(* IEC 61131-3 sources: plc-st-coding-agent/progress/evidence/f14_v10_full_20261113/jobs/custom_deepseek-v4pro (part 5) *)

(* ---- self-hard-02.candidate_02.st ---- *)
(* ENGINEERING_CONTRACT
   - Outputs: phase, elapsed, timeout; initial (0,0,FALSE).
   - Priority: abort > new start edge > run counting (PUB002-006).
   - abortBtn TRUE: phase=9, elapsed/timeout hold previous values. Start edge consumed (PUB003, PUB005-006).
   - New start edge without abort: phase=1, elapsed=0, timeout=FALSE; start scan not counted (PUB004, PUB006).
   - Previous scan running (1 or 2), no abort, no start edge: increment elapsed by 1.
     If elapsed >= maxDuration: timeout=TRUE, phase=3 (timeout priority). Else phase=2 if pv>=setpoint or prevPhase=2, otherwise phase=1 (PUB005-006).
   - Phase 3 complete, phase 9 aborted: freeze elapsed, timeout, phase until new valid start or abort.
   - Unit: elapsed counts scans; maxDuration positive integer scan threshold; comparison >=.
*)
FUNCTION_BLOCK FB
VAR_INPUT
    startBtn : BOOL;
    abortBtn : BOOL;
    setpoint : REAL;
    pv : REAL;
    maxDuration : INT;
END_VAR
VAR_OUTPUT
    elapsed : INT;
    phase : INT;
    timeout : BOOL;
END_VAR
VAR
    prevStartBtn : BOOL := FALSE;
    prevPhase : INT := 0;
    prevElapsed : INT := 0;
    prevTimeout : BOOL := FALSE;
    startEdge : BOOL;
END_VAR

(* Record startBtn rising edge before priority processing; consumed even if abort *)
startEdge := startBtn AND NOT prevStartBtn;

IF abortBtn THEN
    (* Abort highest priority: enter phase 9 and freeze elapsed/timeout *)
    phase := 9;
    elapsed := prevElapsed;
    timeout := prevTimeout;
ELSIF startEdge THEN
    (* New valid start with no abort: reset batch and do not count this scan *)
    phase := 1;
    elapsed := 0;
    timeout := FALSE;
ELSE
    (* No abort and no new start edge *)
    IF (prevPhase = 1) OR (prevPhase = 2) THEN
        (* Running state: count exactly one scan *)
        elapsed := prevElapsed + 1;

        IF elapsed >= maxDuration THEN
            (* Timeout has priority over temperature threshold *)
            timeout := TRUE;
            phase := 3;
        ELSE
            timeout := FALSE;
            IF (prevPhase = 2) OR (pv >= setpoint) THEN
                phase := 2;
            ELSE
                phase := 1;
            END_IF;
        END_IF;
    ELSE
        (* Idle, complete, or aborted: hold state *)
        phase := prevPhase;
        elapsed := prevElapsed;
        timeout := prevTimeout;
    END_IF;
END_IF;

(* Update previous-cycle memory *)
prevStartBtn := startBtn;
prevPhase := phase;
prevElapsed := elapsed;
prevTimeout := timeout;

(* CONTRACT_RULES [] *)
END_FUNCTION_BLOCK

(* ---- self-hard-02.raw_candidate_01.st ---- *)
(* ENGINEERING_CONTRACT
   - phase: 0 idle initial; new start & !abort -> 1; in running, elapsed<maxDuration and (prevPhase=2 or pv>=setpoint) -> 2, else 1; elapsed>=maxDuration -> 3; abort -> 9. Priority abort > start edge > run count (PUB002-006).
   - elapsed: increment exactly once per scan when !abort, !startEdge, prevPhase=1/2; reset 0 on new start; freeze otherwise.
   - timeout: set TRUE exactly when running scan counted reaches maxDuration; reset FALSE on new start; freeze on abort/completion/idle.
   - start rising edge recorded first and consumed even if abort same scan; restart requires release/press.
   - maxDuration positive scan count; comparison >=. Boundaries: counts scan after start not counted.
*)
FUNCTION_BLOCK FB
VAR
    prevStartBtn : BOOL := FALSE;
    prevPhase : INT := 0;
    prevElapsed : INT := 0;
    prevTimeout : BOOL := FALSE;
    startEdge : BOOL;
END_VAR

(* Record startBtn rising edge before priority processing; consumed even if abort *)
startEdge := startBtn AND NOT prevStartBtn;

IF abortBtn THEN
    (* Abort has highest priority: enter phase 9 and freeze elapsed/timeout *)
    phase := 9;
    elapsed := prevElapsed;
    timeout := prevTimeout;
ELSIF startEdge THEN
    (* New valid start with no abort: reset batch and do not count this scan *)
    phase := 1;
    elapsed := 0;
    timeout := FALSE;
ELSE
    (* No abort and no new start edge *)
    IF (prevPhase = 1) OR (prevPhase = 2) THEN
        (* Running state: count exactly one scan *)
        elapsed := prevElapsed + 1;

        IF elapsed >= maxDuration THEN
            (* Timeout has priority over temperature threshold *)
            timeout := TRUE;
            phase := 3;
        ELSE
            timeout := FALSE;
            IF (prevPhase = 2) OR (pv >= setpoint) THEN
                phase := 2;
            ELSE
                phase := 1;
            END_IF;
        END_IF;
    ELSE
        (* Idle, complete, or aborted: hold state *)
        phase := prevPhase;
        elapsed := prevElapsed;
        timeout := prevTimeout;
    END_IF;
END_IF;

(* Update previous-cycle memory *)
prevStartBtn := startBtn;
prevPhase := phase;
prevElapsed := elapsed;
prevTimeout := timeout;

(* CONTRACT_RULES [] *)
END_FUNCTION_BLOCK

(* ---- self-hard-02.raw_candidate_02.st ---- *)
(* ENGINEERING_CONTRACT
   - Outputs: phase, elapsed, timeout; initial (0,0,FALSE).
   - Priority: abort > new start edge > run counting (PUB002-006).
   - abortBtn TRUE: phase=9, elapsed/timeout hold previous values. Start edge consumed (PUB003, PUB005-006).
   - New start edge without abort: phase=1, elapsed=0, timeout=FALSE; start scan not counted (PUB004, PUB006).
   - Previous scan running (1 or 2), no abort, no start edge: increment elapsed by 1.
     If elapsed >= maxDuration: timeout=TRUE, phase=3 (timeout priority). Else phase=2 if pv>=setpoint or prevPhase=2, otherwise phase=1 (PUB005-006).
   - Phase 3 complete, phase 9 aborted: freeze elapsed, timeout, phase until new valid start or abort.
   - Unit: elapsed counts scans; maxDuration positive integer scan threshold; comparison >=.
*)
FUNCTION_BLOCK FB
VAR_INPUT
    startBtn : BOOL;
    abortBtn : BOOL;
    setpoint : REAL;
    pv : REAL;
    maxDuration : INT;
END_VAR
VAR_OUTPUT
    elapsed : INT;
    phase : INT;
    timeout : BOOL;
END_VAR
VAR
    prevStartBtn : BOOL := FALSE;
    prevPhase : INT := 0;
    prevElapsed : INT := 0;
    prevTimeout : BOOL := FALSE;
    startEdge : BOOL;
END_VAR

(* Record startBtn rising edge before priority processing; consumed even if abort *)
startEdge := startBtn AND NOT prevStartBtn;

IF abortBtn THEN
    (* Abort highest priority: enter phase 9 and freeze elapsed/timeout *)
    phase := 9;
    elapsed := prevElapsed;
    timeout := prevTimeout;
ELSIF startEdge THEN
    (* New valid start with no abort: reset batch and do not count this scan *)
    phase := 1;
    elapsed := 0;
    timeout := FALSE;
ELSE
    (* No abort and no new start edge *)
    IF (prevPhase = 1) OR (prevPhase = 2) THEN
        (* Running state: count exactly one scan *)
        elapsed := prevElapsed + 1;

        IF elapsed >= maxDuration THEN
            (* Timeout has priority over temperature threshold *)
            timeout := TRUE;
            phase := 3;
        ELSE
            timeout := FALSE;
            IF (prevPhase = 2) OR (pv >= setpoint) THEN
                phase := 2;
            ELSE
                phase := 1;
            END_IF;
        END_IF;
    ELSE
        (* Idle, complete, or aborted: hold state *)
        phase := prevPhase;
        elapsed := prevElapsed;
        timeout := prevTimeout;
    END_IF;
END_IF;

(* Update previous-cycle memory *)
prevStartBtn := startBtn;
prevPhase := phase;
prevElapsed := elapsed;
prevTimeout := timeout;

(* CONTRACT_RULES [] *)
END_FUNCTION_BLOCK

(* ---- self-hard-03.candidate_01.st ---- *)
(* ENGINEERING_CONTRACT
   Activation: pushEn/popEn rising edges vs stored previous inputs; no repeat while held (PUB001-PUB039).
   Same-scan priority: pop edge is processed first, then push edge; simultaneous full pair frees a slot then appends; simultaneous empty pair adds only new item (PUB001-PUB039).
   Retention: tmp_count is static queue length; fifo[1..tmp_count] stays compact on each scan. No explicit reset; only successful edge actions alter valid queue state (PUB001-PUB039).
   Outputs: count := tmp_count; full := tmp_count = 8; empty := tmp_count = 0; head := fifo[1] when nonempty, else 0 (PUB001-PUB039).
   Bounds: count/INT 0..8; fifo indices 1..8. Invalid tail fifo[tmp_count+1..8] is unspecified and not cleared (PUB001-PUB039).
*)
(* CONTRACT_RULES [] *)
FUNCTION_BLOCK FB
VAR_INPUT
    pushEn : BOOL;
    pushItem : INT;
    popEn : BOOL;
END_VAR
VAR_IN_OUT
    fifo : ARRAY[1..8] OF INT;
END_VAR
VAR_OUTPUT
    count : INT;
    full : BOOL;
    empty : BOOL;
    head : INT;
END_VAR
VAR
    prevPushEn : BOOL := FALSE;
    prevPopEn : BOOL := FALSE;
    tmp_count : INT := 0;
    tmp_pushRise : BOOL;
    tmp_popRise : BOOL;
    tmp_i : INT;
END_VAR

tmp_pushRise := pushEn AND NOT prevPushEn;
tmp_popRise := popEn AND NOT prevPopEn;

IF tmp_popRise THEN
    IF tmp_count > 0 THEN
        IF tmp_count > 1 THEN
            FOR tmp_i := 1 TO tmp_count - 1 DO
                fifo[tmp_i] := fifo[tmp_i + 1];
            END_FOR;
        END_IF;
        tmp_count := tmp_count - 1;
    END_IF;
END_IF;

IF tmp_pushRise THEN
    IF tmp_count < 8 THEN
        tmp_count := tmp_count + 1;
        fifo[tmp_count] := pushItem;
    END_IF;
END_IF;

count := tmp_count;
full := (tmp_count = 8);
empty := (tmp_count = 0);

IF tmp_count > 0 THEN
    head := fifo[1];
ELSE
    head := 0;
END_IF;

prevPushEn := pushEn;
prevPopEn := popEn;

END_FUNCTION_BLOCK

(* ---- self-hard-03.raw_candidate_01.st ---- *)
(* ENGINEERING_CONTRACT
   Activation: pushEn/popEn rising edges vs stored previous inputs; no repeat while held (PUB001-PUB039).
   Same-scan priority: pop edge is processed first, then push edge; simultaneous full pair frees a slot then appends; simultaneous empty pair adds only new item (PUB001-PUB039).
   Retention: tmp_count is static queue length; fifo[1..tmp_count] stays compact on each scan. No explicit reset; only successful edge actions alter valid queue state (PUB001-PUB039).
   Outputs: count := tmp_count; full := tmp_count = 8; empty := tmp_count = 0; head := fifo[1] when nonempty, else 0 (PUB001-PUB039).
   Bounds: count/INT 0..8; fifo indices 1..8. Invalid tail fifo[tmp_count+1..8] is unspecified and not cleared (PUB001-PUB039).
*)
(* CONTRACT_RULES [] *)
FUNCTION_BLOCK FB
VAR_INPUT
    pushEn : BOOL;
    pushItem : INT;
    popEn : BOOL;
END_VAR
VAR_IN_OUT
    fifo : ARRAY[1..8] OF INT;
END_VAR
VAR_OUTPUT
    count : INT;
    full : BOOL;
    empty : BOOL;
    head : INT;
END_VAR
VAR
    prevPushEn : BOOL := FALSE;
    prevPopEn : BOOL := FALSE;
    tmp_count : INT := 0;
    tmp_pushRise : BOOL;
    tmp_popRise : BOOL;
    tmp_i : INT;
END_VAR

tmp_pushRise := pushEn AND NOT prevPushEn;
tmp_popRise := popEn AND NOT prevPopEn;

IF tmp_popRise THEN
    IF tmp_count > 0 THEN
        IF tmp_count > 1 THEN
            FOR tmp_i := 1 TO tmp_count - 1 DO
                fifo[tmp_i] := fifo[tmp_i + 1];
            END_FOR;
        END_IF;
        tmp_count := tmp_count - 1;
    END_IF;
END_IF;

IF tmp_pushRise THEN
    IF tmp_count < 8 THEN
        tmp_count := tmp_count + 1;
        fifo[tmp_count] := pushItem;
    END_IF;
END_IF;

count := tmp_count;
full := (tmp_count = 8);
empty := (tmp_count = 0);

IF tmp_count > 0 THEN
    head := fifo[1];
ELSE
    head := 0;
END_IF;

prevPushEn := pushEn;
prevPopEn := popEn;

END_FUNCTION_BLOCK

(* ---- self-hard-05.candidate_01.st ---- *)
(* ENGINEERING_CONTRACT
   tripLatched: set same-scan on runRequest AND NOT flameOK; held until reset rising edge
                with runRequest=FALSE AND flameOK=FALSE only. Same-scan set/reset mutually exclusive.
   fuelPermit : runRequest AND flameOK AND NOT tripLatched; computed after trip update.
   trimEnable : fuelPermit AND NOT o2Fault.
   airTrim    : trimEnable ? clamp(2.0*(2.0-o2PV), -10.0, 10.0) : 0.0; REAL percent.
   airCommand : fuelPermit ? clamp(baseAir+airTrim, 0.0, 100.0) : 0.0; REAL percent.
   o2Fault    : NOT o2Valid OR o2PV<0.0 OR o2PV>21.0; combinational.
*)
(* CONTRACT_RULES [] *)
FUNCTION_BLOCK FB
VAR_INPUT
    runRequest : BOOL;
    flameOK    : BOOL;
    o2Valid    : BOOL;
    o2PV       : REAL;
    baseAir    : REAL;
    resetBtn   : BOOL;
END_VAR
VAR_OUTPUT
    fuelPermit  : BOOL;
    trimEnable  : BOOL;
    airTrim     : REAL;
    airCommand  : REAL;
    tripLatched : BOOL;
    o2Fault     : BOOL;
END_VAR
VAR
    fbResetEdge     : R_TRIG;
    tmp_resetRising : BOOL;
    tmp_trim        : REAL;
    tmp_cmd         : REAL;
END_VAR

fbResetEdge(CLK := resetBtn);
tmp_resetRising := fbResetEdge.Q;

(* Trip latch: same-scan loss-of-flame set; only valid safe-state reset edge clears. *)
tripLatched := (runRequest AND NOT flameOK)
               OR (tripLatched AND NOT (tmp_resetRising AND NOT runRequest AND NOT flameOK));

(* Oxygen analyzer fault and permits. *)
o2Fault := (NOT o2Valid) OR (o2PV < 0.0) OR (o2PV > 21.0);
fuelPermit := runRequest AND flameOK AND NOT tripLatched;
trimEnable := fuelPermit AND NOT o2Fault;

(* Oxygen trim with +/-10 percent output clamp. *)
IF trimEnable THEN
    tmp_trim := 2.0 * (2.0 - o2PV);
    IF tmp_trim < -10.0 THEN
        tmp_trim := -10.0;
    ELSIF tmp_trim > 10.0 THEN
        tmp_trim := 10.0;
    END_IF;
    airTrim := tmp_trim;
ELSE
    airTrim := 0.0;
END_IF;

(* Final air command with 0..100 percent output clamp. *)
IF fuelPermit THEN
    tmp_cmd := baseAir + airTrim;
    IF tmp_cmd < 0.0 THEN
        tmp_cmd := 0.0;
    ELSIF tmp_cmd > 100.0 THEN
        tmp_cmd := 100.0;
    END_IF;
    airCommand := tmp_cmd;
ELSE
    airCommand := 0.0;
END_IF;

END_FUNCTION_BLOCK

(* ---- self-hard-05.raw_candidate_01.st ---- *)
(* ENGINEERING_CONTRACT
   tripLatched: set same-scan on runRequest AND NOT flameOK; held until reset rising edge
                with runRequest=FALSE AND flameOK=FALSE only. Same-scan set/reset mutually exclusive.
   fuelPermit : runRequest AND flameOK AND NOT tripLatched; computed after trip update.
   trimEnable : fuelPermit AND NOT o2Fault.
   airTrim    : trimEnable ? clamp(2.0*(2.0-o2PV), -10.0, 10.0) : 0.0; REAL percent.
   airCommand : fuelPermit ? clamp(baseAir+airTrim, 0.0, 100.0) : 0.0; REAL percent.
   o2Fault    : NOT o2Valid OR o2PV<0.0 OR o2PV>21.0; combinational.
*)
(* CONTRACT_RULES [] *)
FUNCTION_BLOCK FB
VAR_INPUT
    runRequest : BOOL;
    flameOK    : BOOL;
    o2Valid    : BOOL;
    o2PV       : REAL;
    baseAir    : REAL;
    resetBtn   : BOOL;
END_VAR
VAR_OUTPUT
    fuelPermit  : BOOL;
    trimEnable  : BOOL;
    airTrim     : REAL;
    airCommand  : REAL;
    tripLatched : BOOL;
    o2Fault     : BOOL;
END_VAR
VAR
    fbResetEdge     : R_TRIG;
    tmp_resetRising : BOOL;
    tmp_trim        : REAL;
    tmp_cmd         : REAL;
END_VAR

fbResetEdge(CLK := resetBtn);
tmp_resetRising := fbResetEdge.Q;

(* Trip latch: same-scan loss-of-flame set; only valid safe-state reset edge clears. *)
tripLatched := (runRequest AND NOT flameOK)
               OR (tripLatched AND NOT (tmp_resetRising AND NOT runRequest AND NOT flameOK));

(* Oxygen analyzer fault and permits. *)
o2Fault := (NOT o2Valid) OR (o2PV < 0.0) OR (o2PV > 21.0);
fuelPermit := runRequest AND flameOK AND NOT tripLatched;
trimEnable := fuelPermit AND NOT o2Fault;

(* Oxygen trim with +/-10 percent output clamp. *)
IF trimEnable THEN
    tmp_trim := 2.0 * (2.0 - o2PV);
    IF tmp_trim < -10.0 THEN
        tmp_trim := -10.0;
    ELSIF tmp_trim > 10.0 THEN
        tmp_trim := 10.0;
    END_IF;
    airTrim := tmp_trim;
ELSE
    airTrim := 0.0;
END_IF;

(* Final air command with 0..100 percent output clamp. *)
IF fuelPermit THEN
    tmp_cmd := baseAir + airTrim;
    IF tmp_cmd < 0.0 THEN
        tmp_cmd := 0.0;
    ELSIF tmp_cmd > 100.0 THEN
        tmp_cmd := 100.0;
    END_IF;
    airCommand := tmp_cmd;
ELSE
    airCommand := 0.0;
END_IF;

END_FUNCTION_BLOCK

(* ---- self-hard-06.candidate_01.st ---- *)
(* ENGINEERING_CONTRACT
   - tripLatched: set same scan by run & (!valid | P>=4500) PUB002/PUB006; holds until legal reset edge.
     Legal reset: rising reset & !run & valid & P<=4200 PUB003. Illegal reset does not clear PUB012/PUB013.
   - currentCauseMask: recomputed each scan; allowed 0/1/2/4/6/8 PUB008,N10-S15.
     bit0=invalid; bit1 requires 3 consecutive full stuck scans PUB010,N10-S11; bit2 inclusive flow; bit3=8 when no located bit under overpressure.
   - latchedCauseMask: OR-accumulates currentCauseMask while tripLatched true; cleared when not tripped or legal reset PUB011,N10-S18.
   - fuelPermit = run & !trip; diagnosticActive = current<>0 PUB007.
   - stuck counter zeroes on any non-full scan: !run, !valid, P<4500, or valve condition false PUB010.
   - units: kPa, t/h, %; boundaries inclusive. Same-scan trip and cause are emitted together.
*)
(* CONTRACT_RULES [] *)
FUNCTION_BLOCK FB
VAR_INPUT
    runRequest: BOOL;
    pressure: REAL;
    pressureValid: BOOL;
    fuelFlow: REAL;
    steamFlow: REAL;
    outletCmd: INT;
    outletFeedback: INT;
    resetBtn: BOOL;
END_VAR
VAR_OUTPUT
    tripLatched: BOOL;
    fuelPermit: BOOL;
    currentCauseMask: WORD;
    latchedCauseMask: WORD;
    diagnosticActive: BOOL;
END_VAR
VAR
    prev_reset_btn: BOOL := FALSE;
    prev_trip_state: BOOL := FALSE;
    stuck_count: INT := 0;
    latched_state: WORD := WORD#16#0000;
    tmp_rising_reset: BOOL;
    tmp_legal_reset: BOOL;
    tmp_stuck_condition: BOOL;
    tmp_bit1: BOOL;
    tmp_bit2: BOOL;
    tmp_trip_condition: BOOL;
    tmp_trip_state: BOOL;
END_VAR

(* Update stuck-valve consecutive-scan counter *)
tmp_stuck_condition := runRequest AND pressureValid AND (pressure >= 4500.0)
                       AND (outletCmd >= 50) AND (outletFeedback <= 10);

IF tmp_stuck_condition THEN
    IF stuck_count < 3 THEN
        stuck_count := stuck_count + 1;
    END_IF;
ELSE
    stuck_count := 0;
END_IF;

(* Compute current cause mask *)
currentCauseMask := WORD#16#0000;

IF NOT runRequest THEN
    currentCauseMask := WORD#16#0000;
ELSIF NOT pressureValid THEN
    currentCauseMask := WORD#16#0001; (* bit0: transmitter invalid *)
ELSE
    IF pressure >= 4500.0 THEN
        tmp_bit1 := stuck_count >= 3;
        tmp_bit2 := (fuelFlow >= 4.0) AND (steamFlow <= 10.0);

        IF tmp_bit1 THEN
            currentCauseMask := currentCauseMask OR WORD#16#0002; (* bit1: valve stuck *)
        END_IF;
        IF tmp_bit2 THEN
            currentCauseMask := currentCauseMask OR WORD#16#0004; (* bit2: combustion excess *)
        END_IF;
        IF currentCauseMask = WORD#16#0000 THEN
            currentCauseMask := WORD#16#0008; (* bit3: not located *)
        END_IF;
    ELSE
        currentCauseMask := WORD#16#0000;
    END_IF;
END_IF;

(* Trip latch state *)
tmp_rising_reset := resetBtn AND NOT prev_reset_btn;
tmp_legal_reset := tmp_rising_reset AND (NOT runRequest) AND pressureValid AND (pressure <= 4200.0);

tmp_trip_condition := runRequest AND ((NOT pressureValid) OR (pressureValid AND (pressure >= 4500.0)));
tmp_trip_state := tmp_trip_condition OR (prev_trip_state AND NOT tmp_legal_reset);
tripLatched := tmp_trip_state;

(* Latched footprint accumulation / clear *)
IF tmp_trip_state THEN
    latched_state := (latched_state OR currentCauseMask) AND WORD#16#000F;
ELSE
    latched_state := WORD#16#0000;
END_IF;
latchedCauseMask := latched_state;

(* Derived outputs *)
fuelPermit := runRequest AND NOT tripLatched;
diagnosticActive := currentCauseMask <> WORD#16#0000;

(* Remember previous-scan values for next call *)
prev_reset_btn := resetBtn;
prev_trip_state := tmp_trip_state;

END_FUNCTION_BLOCK

(* ---- self-hard-06.raw_candidate_01.st ---- *)
(* ENGINEERING_CONTRACT
   - tripLatched: set same scan by run & (!valid | P>=4500) PUB002/PUB006; holds until legal reset edge.
     Legal reset: rising reset & !run & valid & P<=4200 PUB003. Illegal reset does not clear PUB012/PUB013.
   - currentCauseMask: recomputed each scan; allowed 0/1/2/4/6/8 PUB008,N10-S15.
     bit0=invalid; bit1 requires 3 consecutive full stuck scans PUB010,N10-S11; bit2 inclusive flow; bit3=8 when no located bit under overpressure.
   - latchedCauseMask: OR-accumulates currentCauseMask while tripLatched true; cleared when not tripped or legal reset PUB011,N10-S18.
   - fuelPermit = run & !trip; diagnosticActive = current<>0 PUB007.
   - stuck counter zeroes on any non-full scan: !run, !valid, P<4500, or valve condition false PUB010.
   - units: kPa, t/h, %; boundaries inclusive. Same-scan trip and cause are emitted together.
*)
(* CONTRACT_RULES [] *)
FUNCTION_BLOCK FB
VAR_INPUT
    runRequest: BOOL;
    pressure: REAL;
    pressureValid: BOOL;
    fuelFlow: REAL;
    steamFlow: REAL;
    outletCmd: INT;
    outletFeedback: INT;
    resetBtn: BOOL;
END_VAR
VAR_OUTPUT
    tripLatched: BOOL;
    fuelPermit: BOOL;
    currentCauseMask: WORD;
    latchedCauseMask: WORD;
    diagnosticActive: BOOL;
END_VAR
VAR
    prev_reset_btn: BOOL := FALSE;
    prev_trip_state: BOOL := FALSE;
    stuck_count: INT := 0;
    latched_state: WORD := WORD#16#0000;
    tmp_rising_reset: BOOL;
    tmp_legal_reset: BOOL;
    tmp_stuck_condition: BOOL;
    tmp_bit1: BOOL;
    tmp_bit2: BOOL;
    tmp_trip_condition: BOOL;
    tmp_trip_state: BOOL;
END_VAR

(* Update stuck-valve consecutive-scan counter *)
tmp_stuck_condition := runRequest AND pressureValid AND (pressure >= 4500.0)
                       AND (outletCmd >= 50) AND (outletFeedback <= 10);

IF tmp_stuck_condition THEN
    IF stuck_count < 3 THEN
        stuck_count := stuck_count + 1;
    END_IF;
ELSE
    stuck_count := 0;
END_IF;

(* Compute current cause mask *)
currentCauseMask := WORD#16#0000;

IF NOT runRequest THEN
    currentCauseMask := WORD#16#0000;
ELSIF NOT pressureValid THEN
    currentCauseMask := WORD#16#0001; (* bit0: transmitter invalid *)
ELSE
    IF pressure >= 4500.0 THEN
        tmp_bit1 := stuck_count >= 3;
        tmp_bit2 := (fuelFlow >= 4.0) AND (steamFlow <= 10.0);

        IF tmp_bit1 THEN
            currentCauseMask := currentCauseMask OR WORD#16#0002; (* bit1: valve stuck *)
        END_IF;
        IF tmp_bit2 THEN
            currentCauseMask := currentCauseMask OR WORD#16#0004; (* bit2: combustion excess *)
        END_IF;
        IF currentCauseMask = WORD#16#0000 THEN
            currentCauseMask := WORD#16#0008; (* bit3: not located *)
        END_IF;
    ELSE
        currentCauseMask := WORD#16#0000;
    END_IF;
END_IF;

(* Trip latch state *)
tmp_rising_reset := resetBtn AND NOT prev_reset_btn;
tmp_legal_reset := tmp_rising_reset AND (NOT runRequest) AND pressureValid AND (pressure <= 4200.0);

tmp_trip_condition := runRequest AND ((NOT pressureValid) OR (pressureValid AND (pressure >= 4500.0)));
tmp_trip_state := tmp_trip_condition OR (prev_trip_state AND NOT tmp_legal_reset);
tripLatched := tmp_trip_state;

(* Latched footprint accumulation / clear *)
IF tmp_trip_state THEN
    latched_state := (latched_state OR currentCauseMask) AND WORD#16#000F;
ELSE
    latched_state := WORD#16#0000;
END_IF;
latchedCauseMask := latched_state;

(* Derived outputs *)
fuelPermit := runRequest AND NOT tripLatched;
diagnosticActive := currentCauseMask <> WORD#16#0000;

(* Remember previous-scan values for next call *)
prev_reset_btn := resetBtn;
prev_trip_state := tmp_trip_state;

END_FUNCTION_BLOCK

(* ---- self-medium-01.candidate_01.st ---- *)
TYPE ST_Recipe :
STRUCT
    recipeID : INT;
    totalRatio : REAL;
    temperature : REAL;
END_STRUCT
END_TYPE;

(* ENGINEERING_CONTRACT
   valid/loadedID activate only on loadCmd rising edge with running=FALSE (PUB003/PUB007/PUB010).
   Legal slot check 1..8 precedes any array access; out-of-range is not indexed (PUB006/S5).
   Candidate = recipeID<>0 AND totalRatio in [99.0,101.0] AND temperature in [30.0,180.0] (PUB008/N10-S7).
   Accepted invalid edge clears valid=FALSE and loadedID=0; valid edge loads selected recipeID (PUB009/N10-S8/S1).
   running=TRUE overrides any load edge and holds previous valid/loadedID (PUB010/N10-S4/N10-S9).
   No rising edge holds previous outputs (S6/S9).
   Units/bounds: REAL closed intervals; no timing; selSlot dimensionless.
   Conflict note: F13-S1 prose says empty-slot must not change ID, but formal S1/N10-S8/req5 require clear; clear is implemented.
*)

(* CONTRACT_RULES [] *)

FUNCTION_BLOCK FB
VAR_INPUT
    recipe : ARRAY[1..8] OF ST_Recipe;
    selSlot : INT;
    loadCmd : BOOL;
    running : BOOL;
END_VAR
VAR_OUTPUT
    valid : BOOL;
    loadedID : INT;
END_VAR
VAR
    tmp_prevLoadCmd : BOOL := FALSE;
    tmp_validState : BOOL := FALSE;
    tmp_loadedIDState : INT := 0;
    tmp_edge : BOOL;
    tmp_slotLegal : BOOL;
    tmp_candidateValid : BOOL;
    tmp_isNonEmpty : BOOL;
    tmp_ratioOk : BOOL;
    tmp_tempOk : BOOL;
    tmp_recipeId : INT;
    tmp_totalRatio : REAL;
    tmp_temperature : REAL;
END_VAR

tmp_edge := loadCmd AND NOT tmp_prevLoadCmd;

IF (NOT running) AND tmp_edge THEN
    tmp_slotLegal := (selSlot >= 1) AND (selSlot <= 8);
    IF tmp_slotLegal THEN
        tmp_recipeId := recipe[selSlot].recipeID;
        tmp_totalRatio := recipe[selSlot].totalRatio;
        tmp_temperature := recipe[selSlot].temperature;

        tmp_isNonEmpty := (tmp_recipeId <> 0);
        tmp_ratioOk := (tmp_totalRatio >= 99.0) AND (tmp_totalRatio <= 101.0);
        tmp_tempOk := (tmp_temperature >= 30.0) AND (tmp_temperature <= 180.0);
        tmp_candidateValid := tmp_isNonEmpty AND tmp_ratioOk AND tmp_tempOk;

        tmp_validState := tmp_candidateValid;
        IF tmp_candidateValid THEN
            tmp_loadedIDState := tmp_recipeId;
        ELSE
            tmp_loadedIDState := 0;
        END_IF;
    ELSE
        tmp_validState := FALSE;
        tmp_loadedIDState := 0;
    END_IF;
END_IF;

valid := tmp_validState;
loadedID := tmp_loadedIDState;
tmp_prevLoadCmd := loadCmd;

END_FUNCTION_BLOCK

(* ---- self-medium-01.raw_candidate_01.st ---- *)
TYPE ST_Recipe :
STRUCT
    recipeID : INT;
    totalRatio : REAL;
    temperature : REAL;
END_STRUCT
END_TYPE

(* ENGINEERING_CONTRACT
   valid/loadedID activate only on loadCmd rising edge with running=FALSE (PUB003/PUB007/PUB010).
   Legal slot check 1..8 precedes any array access; out-of-range is not indexed (PUB006/S5).
   Candidate = recipeID<>0 AND totalRatio in [99.0,101.0] AND temperature in [30.0,180.0] (PUB008/N10-S7).
   Accepted invalid edge clears valid=FALSE and loadedID=0; valid edge loads selected recipeID (PUB009/N10-S8/S1).
   running=TRUE overrides any load edge and holds previous valid/loadedID (PUB010/N10-S4/N10-S9).
   No rising edge holds previous outputs (S6/S9).
   Units/bounds: REAL closed intervals; no timing; selSlot dimensionless.
   Conflict note: F13-S1 prose says empty-slot must not change ID, but formal S1/N10-S8/req5 require clear; clear is implemented.
*)

(* CONTRACT_RULES [] *)

FUNCTION_BLOCK FB
VAR_INPUT
    recipe : ARRAY[1..8] OF ST_Recipe;
    selSlot : INT;
    loadCmd : BOOL;
    running : BOOL;
END_VAR
VAR_OUTPUT
    valid : BOOL;
    loadedID : INT;
END_VAR
VAR
    tmp_prevLoadCmd : BOOL := FALSE;
    tmp_validState : BOOL := FALSE;
    tmp_loadedIDState : INT := 0;
    tmp_edge : BOOL;
    tmp_slotLegal : BOOL;
    tmp_candidateValid : BOOL;
    tmp_isNonEmpty : BOOL;
    tmp_ratioOk : BOOL;
    tmp_tempOk : BOOL;
    tmp_recipeId : INT;
    tmp_totalRatio : REAL;
    tmp_temperature : REAL;
END_VAR

tmp_edge := loadCmd AND NOT tmp_prevLoadCmd;

IF (NOT running) AND tmp_edge THEN
    tmp_slotLegal := (selSlot >= 1) AND (selSlot <= 8);
    IF tmp_slotLegal THEN
        tmp_recipeId := recipe[selSlot].recipeID;
        tmp_totalRatio := recipe[selSlot].totalRatio;
        tmp_temperature := recipe[selSlot].temperature;

        tmp_isNonEmpty := (tmp_recipeId <> 0);
        tmp_ratioOk := (tmp_totalRatio >= 99.0) AND (tmp_totalRatio <= 101.0);
        tmp_tempOk := (tmp_temperature >= 30.0) AND (tmp_temperature <= 180.0);
        tmp_candidateValid := tmp_isNonEmpty AND tmp_ratioOk AND tmp_tempOk;

        tmp_validState := tmp_candidateValid;
        IF tmp_candidateValid THEN
            tmp_loadedIDState := tmp_recipeId;
        ELSE
            tmp_loadedIDState := 0;
        END_IF;
    ELSE
        tmp_validState := FALSE;
        tmp_loadedIDState := 0;
    END_IF;
END_IF;

valid := tmp_validState;
loadedID := tmp_loadedIDState;
tmp_prevLoadCmd := loadCmd;

END_FUNCTION_BLOCK

(* ---- self-medium-02.candidate_01.st ---- *)
FUNCTION_BLOCK FB
VAR_INPUT
    enable : BOOL;
    rawValue : REAL;
END_VAR
VAR_OUTPUT
    filteredValue : REAL;
    windowFull : BOOL;
    sampleCount : INT;
END_VAR
VAR
    local_data : ARRAY[0..7] OF REAL;
    local_count : INT := 0;
    local_writeIdx : INT := 0;
    local_sum : REAL;
    local_idx : INT;
    local_filtered : REAL := 0.0;
END_VAR

(* ENGINEERING_CONTRACT
  [PUB001-PUB003] enable TRUE: insert rawValue into 8-slot FIFO.
  [PUB004-PUB008] count=min(8,prev+1); unfilled slots ignored.
  [PUB009-PUB012] full: replace oldest slot and rotate write index.
  [PUB013-PUB016] sampleCount=count 0..8; windowFull=(count=8).
  [PUB017-PUB020] enable FALSE: clear history, count=0, full=FALSE,
      filteredValue held from last computation.
  [S1-S7] average over first count slots; boundaries strict; output at end.
*)

(* CONTRACT_RULES [] *)

IF enable THEN
    IF local_count < 8 THEN
        local_data[local_count] := rawValue;
        local_count := local_count + 1;
        local_writeIdx := local_count MOD 8;
    ELSE
        local_data[local_writeIdx] := rawValue;
        local_writeIdx := (local_writeIdx + 1) MOD 8;
    END_IF;

    sampleCount := local_count;
    windowFull := (local_count = 8);

    local_sum := 0.0;
    FOR local_idx := 0 TO local_count - 1 DO
        local_sum := local_sum + local_data[local_idx];
    END_FOR;

    local_filtered := local_sum / INT_TO_REAL(local_count);
    filteredValue := local_filtered;
ELSE
    local_count := 0;
    local_writeIdx := 0;
    sampleCount := 0;
    windowFull := FALSE;

    FOR local_idx := 0 TO 7 DO
        local_data[local_idx] := 0.0;
    END_FOR;

    filteredValue := local_filtered;
END_IF;
END_FUNCTION_BLOCK

(* ---- self-medium-02.raw_candidate_01.st ---- *)
FUNCTION_BLOCK FB
VAR_INPUT
    enable : BOOL;
    rawValue : REAL;
END_VAR
VAR_OUTPUT
    filteredValue : REAL;
    windowFull : BOOL;
    sampleCount : INT;
END_VAR
VAR
    local_data : ARRAY[0..7] OF REAL;
    local_count : INT := 0;
    local_writeIdx : INT := 0;
    local_sum : REAL;
    local_idx : INT;
    local_filtered : REAL := 0.0;
END_VAR

(* ENGINEERING_CONTRACT
  [PUB001-PUB003] enable TRUE: insert rawValue into 8-slot FIFO.
  [PUB004-PUB008] count=min(8,prev+1); unfilled slots ignored.
  [PUB009-PUB012] full: replace oldest slot and rotate write index.
  [PUB013-PUB016] sampleCount=count 0..8; windowFull=(count=8).
  [PUB017-PUB020] enable FALSE: clear history, count=0, full=FALSE,
      filteredValue held from last computation.
  [S1-S7] average over first count slots; boundaries strict; output at end.
*)

(* CONTRACT_RULES [] *)

IF enable THEN
    IF local_count < 8 THEN
        local_data[local_count] := rawValue;
        local_count := local_count + 1;
        local_writeIdx := local_count MOD 8;
    ELSE
        local_data[local_writeIdx] := rawValue;
        local_writeIdx := (local_writeIdx + 1) MOD 8;
    END_IF;

    sampleCount := local_count;
    windowFull := (local_count = 8);

    local_sum := 0.0;
    FOR local_idx := 0 TO local_count - 1 DO
        local_sum := local_sum + local_data[local_idx];
    END_FOR;

    local_filtered := local_sum / INT_TO_REAL(local_count);
    filteredValue := local_filtered;
ELSE
    local_count := 0;
    local_writeIdx := 0;
    sampleCount := 0;
    windowFull := FALSE;

    FOR local_idx := 0 TO 7 DO
        local_data[local_idx] := 0.0;
    END_FOR;

    filteredValue := local_filtered;
END_IF;
END_FUNCTION_BLOCK

(* ---- self-medium-03.candidate_01.st ---- *)
(* ENGINEERING_CONTRACT
   state IDLE/OPENING/CLOSING/FAULT retained in FB; initial IDLE, all previous inputs/outputs FALSE.
   motorUp: activates on IDLE legal open edge, holds while no obstacle and no openLimit; stops at limit/obstacle/fault; mutually exclusive with down.
   motorDown: symmetric close handling, holds while no obstacle and no closeLimit; mutually exclusive with up.
   errorFlag: set by obstacle any scan; latched until bothBTN rising edge and no obstacle; obstacle overrides reset; reset scan motors off, state IDLE.
   prev* memory updated after outputs; BOOL units, initial prev FALSE.
*)
(* CONTRACT_RULES [] *)
FUNCTION_BLOCK FB
VAR
    state : INT := 0; (* 0=IDLE, 1=OPENING, 2=CLOSING, 3=FAULT *)
    prevOpenBtn : BOOL := FALSE;
    prevCloseBtn : BOOL := FALSE;
    prevBothBtn : BOOL := FALSE;
    prevMotorUp : BOOL := FALSE;
    prevMotorDown : BOOL := FALSE;
    prevErrorFlag : BOOL := FALSE;
    prevObstacle : BOOL := FALSE;
    risingOpen : BOOL;
    risingClose : BOOL;
    risingBoth : BOOL;
END_VAR

risingOpen := openBtn AND (NOT prevOpenBtn);
risingClose := closeBtn AND (NOT prevCloseBtn);
risingBoth := (openBtn AND closeBtn) AND (NOT prevBothBtn);

motorUp := (NOT obstacle) AND (NOT openLimit) AND
           (prevMotorUp OR
            ((NOT prevMotorUp) AND (NOT prevMotorDown) AND
             (NOT prevErrorFlag) AND risingOpen AND (NOT closeBtn)));

motorDown := (NOT obstacle) AND (NOT closeLimit) AND
             (prevMotorDown OR
              ((NOT prevMotorUp) AND (NOT prevMotorDown) AND
               (NOT prevErrorFlag) AND risingClose AND (NOT openBtn)));

errorFlag := obstacle OR (prevErrorFlag AND (NOT risingBoth));

IF obstacle THEN
    state := 3;
ELSIF state = 3 THEN
    IF risingBoth THEN
        state := 0;
    ELSE
        state := 3;
    END_IF;
ELSE
    IF motorUp THEN
        state := 1;
    ELSIF motorDown THEN
        state := 2;
    ELSE
        state := 0;
    END_IF;
END_IF;

prevOpenBtn := openBtn;
prevCloseBtn := closeBtn;
prevBothBtn := openBtn AND closeBtn;
prevMotorUp := motorUp;
prevMotorDown := motorDown;
prevErrorFlag := errorFlag;
prevObstacle := obstacle;

END_FUNCTION_BLOCK

(* ---- self-medium-03.candidate_02.st ---- *)
(* ENGINEERING_CONTRACT
   State IDLE/OPENING/CLOSING/FAULT retained in FB; initial IDLE, all previous inputs/outputs FALSE.
   motorUp: activates on IDLE legal open edge, holds while no obstacle and no openLimit; stops at limit/obstacle/fault.
   motorDown: symmetric close handling, holds while no obstacle and no closeLimit.
   errorFlag: set by obstacle any scan; latched until bothBTN rising edge and no obstacle; obstacle overrides reset.
   prev* memory updated after outputs; BOOL units, initial prev FALSE.
*)
(* CONTRACT_RULES [] *)
FUNCTION_BLOCK FB
VAR_INPUT
    openBtn : BOOL;
    closeBtn : BOOL;
    openLimit : BOOL;
    closeLimit : BOOL;
    obstacle : BOOL;
END_VAR
VAR_OUTPUT
    motorUp : BOOL;
    motorDown : BOOL;
    errorFlag : BOOL;
END_VAR
VAR
    state : INT := 0; (* 0=IDLE, 1=OPENING, 2=CLOSING, 3=FAULT *)
    prevOpenBtn : BOOL := FALSE;
    prevCloseBtn : BOOL := FALSE;
    prevBothBtn : BOOL := FALSE;
    prevMotorUp : BOOL := FALSE;
    prevMotorDown : BOOL := FALSE;
    prevErrorFlag : BOOL := FALSE;
    prevObstacle : BOOL := FALSE;
    risingOpen : BOOL;
    risingClose : BOOL;
    risingBoth : BOOL;
END_VAR

risingOpen := openBtn AND (NOT prevOpenBtn);
risingClose := closeBtn AND (NOT prevCloseBtn);
risingBoth := (openBtn AND closeBtn) AND (NOT prevBothBtn);

motorUp := (NOT obstacle) AND (NOT openLimit) AND
           (prevMotorUp OR
            ((NOT prevMotorUp) AND (NOT prevMotorDown) AND
             (NOT prevErrorFlag) AND risingOpen AND (NOT closeBtn)));

motorDown := (NOT obstacle) AND (NOT closeLimit) AND
             (prevMotorDown OR
              ((NOT prevMotorUp) AND (NOT prevMotorDown) AND
               (NOT prevErrorFlag) AND risingClose AND (NOT openBtn)));

errorFlag := obstacle OR (prevErrorFlag AND (NOT risingBoth));

IF obstacle THEN
    state := 3;
ELSIF state = 3 THEN
    IF risingBoth THEN
        state := 0;
    ELSE
        state := 3;
    END_IF;
ELSE
    IF motorUp THEN
        state := 1;
    ELSIF motorDown THEN
        state := 2;
    ELSE
        state := 0;
    END_IF;
END_IF;

prevOpenBtn := openBtn;
prevCloseBtn := closeBtn;
prevBothBtn := openBtn AND closeBtn;
prevMotorUp := motorUp;
prevMotorDown := motorDown;
prevErrorFlag := errorFlag;
prevObstacle := obstacle;

END_FUNCTION_BLOCK

(* ---- self-medium-03.raw_candidate_01.st ---- *)
(* ENGINEERING_CONTRACT
   state IDLE/OPENING/CLOSING/FAULT retained in FB; initial IDLE, all previous inputs/outputs FALSE.
   motorUp: activates on IDLE legal open edge, holds while no obstacle and no openLimit; stops at limit/obstacle/fault; mutually exclusive with down.
   motorDown: symmetric close handling, holds while no obstacle and no closeLimit; mutually exclusive with up.
   errorFlag: set by obstacle any scan; latched until bothBTN rising edge and no obstacle; obstacle overrides reset; reset scan motors off, state IDLE.
   prev* memory updated after outputs; BOOL units, initial prev FALSE.
*)
(* CONTRACT_RULES [] *)
FUNCTION_BLOCK FB
VAR
    state : INT := 0; (* 0=IDLE, 1=OPENING, 2=CLOSING, 3=FAULT *)
    prevOpenBtn : BOOL := FALSE;
    prevCloseBtn : BOOL := FALSE;
    prevBothBtn : BOOL := FALSE;
    prevMotorUp : BOOL := FALSE;
    prevMotorDown : BOOL := FALSE;
    prevErrorFlag : BOOL := FALSE;
    prevObstacle : BOOL := FALSE;
    risingOpen : BOOL;
    risingClose : BOOL;
    risingBoth : BOOL;
END_VAR

risingOpen := openBtn AND (NOT prevOpenBtn);
risingClose := closeBtn AND (NOT prevCloseBtn);
risingBoth := (openBtn AND closeBtn) AND (NOT prevBothBtn);

motorUp := (NOT obstacle) AND (NOT openLimit) AND
           (prevMotorUp OR
            ((NOT prevMotorUp) AND (NOT prevMotorDown) AND
             (NOT prevErrorFlag) AND risingOpen AND (NOT closeBtn)));

motorDown := (NOT obstacle) AND (NOT closeLimit) AND
             (prevMotorDown OR
              ((NOT prevMotorUp) AND (NOT prevMotorDown) AND
               (NOT prevErrorFlag) AND risingClose AND (NOT openBtn)));

errorFlag := obstacle OR (prevErrorFlag AND (NOT risingBoth));

IF obstacle THEN
    state := 3;
ELSIF state = 3 THEN
    IF risingBoth THEN
        state := 0;
    ELSE
        state := 3;
    END_IF;
ELSE
    IF motorUp THEN
        state := 1;
    ELSIF motorDown THEN
        state := 2;
    ELSE
        state := 0;
    END_IF;
END_IF;

prevOpenBtn := openBtn;
prevCloseBtn := closeBtn;
prevBothBtn := openBtn AND closeBtn;
prevMotorUp := motorUp;
prevMotorDown := motorDown;
prevErrorFlag := errorFlag;
prevObstacle := obstacle;

END_FUNCTION_BLOCK

(* ---- self-medium-03.raw_candidate_02.st ---- *)
(* ENGINEERING_CONTRACT
   State IDLE/OPENING/CLOSING/FAULT retained in FB; initial IDLE, all previous inputs/outputs FALSE.
   motorUp: activates on IDLE legal open edge, holds while no obstacle and no openLimit; stops at limit/obstacle/fault.
   motorDown: symmetric close handling, holds while no obstacle and no closeLimit.
   errorFlag: set by obstacle any scan; latched until bothBTN rising edge and no obstacle; obstacle overrides reset.
   prev* memory updated after outputs; BOOL units, initial prev FALSE.
*)
(* CONTRACT_RULES [] *)
FUNCTION_BLOCK FB
VAR_INPUT
    openBtn : BOOL;
    closeBtn : BOOL;
    openLimit : BOOL;
    closeLimit : BOOL;
    obstacle : BOOL;
END_VAR
VAR_OUTPUT
    motorUp : BOOL;
    motorDown : BOOL;
    errorFlag : BOOL;
END_VAR
VAR
    state : INT := 0; (* 0=IDLE, 1=OPENING, 2=CLOSING, 3=FAULT *)
    prevOpenBtn : BOOL := FALSE;
    prevCloseBtn : BOOL := FALSE;
    prevBothBtn : BOOL := FALSE;
    prevMotorUp : BOOL := FALSE;
    prevMotorDown : BOOL := FALSE;
    prevErrorFlag : BOOL := FALSE;
    prevObstacle : BOOL := FALSE;
    risingOpen : BOOL;
    risingClose : BOOL;
    risingBoth : BOOL;
END_VAR

risingOpen := openBtn AND (NOT prevOpenBtn);
risingClose := closeBtn AND (NOT prevCloseBtn);
risingBoth := (openBtn AND closeBtn) AND (NOT prevBothBtn);

motorUp := (NOT obstacle) AND (NOT openLimit) AND
           (prevMotorUp OR
            ((NOT prevMotorUp) AND (NOT prevMotorDown) AND
             (NOT prevErrorFlag) AND risingOpen AND (NOT closeBtn)));

motorDown := (NOT obstacle) AND (NOT closeLimit) AND
             (prevMotorDown OR
              ((NOT prevMotorUp) AND (NOT prevMotorDown) AND
               (NOT prevErrorFlag) AND risingClose AND (NOT openBtn)));

errorFlag := obstacle OR (prevErrorFlag AND (NOT risingBoth));

IF obstacle THEN
    state := 3;
ELSIF state = 3 THEN
    IF risingBoth THEN
        state := 0;
    ELSE
        state := 3;
    END_IF;
ELSE
    IF motorUp THEN
        state := 1;
    ELSIF motorDown THEN
        state := 2;
    ELSE
        state := 0;
    END_IF;
END_IF;

prevOpenBtn := openBtn;
prevCloseBtn := closeBtn;
prevBothBtn := openBtn AND closeBtn;
prevMotorUp := motorUp;
prevMotorDown := motorDown;
prevErrorFlag := errorFlag;
prevObstacle := obstacle;

END_FUNCTION_BLOCK

(* ---- self-medium-04.candidate_01.st ---- *)
FUNCTION_BLOCK FB
VAR_INPUT
    startBtn : BOOL;
    resetBtn : BOOL;
    doneSensor : BOOL;
    targetVol : REAL;
    flowVol : REAL;
END_VAR
VAR_OUTPUT
    valveOpen : BOOL;
    fillsToday : INT;
END_VAR
VAR
    start_prev : BOOL := FALSE;
    reset_prev : BOOL := FALSE;
    pendingConfirm : BOOL := FALSE;
    local_accumVol : REAL := 0.0;
    local_start_rise : BOOL;
    local_reset_rise : BOOL;
END_VAR

(* ENGINEERING_CONTRACT
valveOpen: set on start_rise while previous output closed; hold while accumulated volume < targetVol;
            reset_rise priority closes immediately (S2,S5,S7,S8,S9).
pendingConfirm: set when accumulated volume reaches targetVol and valve closes; cleared by reset, new start,
            or confirmation after doneSensor = TRUE (Step4,S10,S13,S14).
fillsToday: +1 on pendingConfirm AND doneSensor, saturating at INT#32767; reset_rise sets 0;
            monotonic except reset (S1,S3,S4,S6,S14).
accumVol: REAL, mL; targetVol and flowVol REAL, mL; comparison uses >=.
*)
(* CONTRACT_RULES [] *)

local_start_rise := startBtn AND NOT start_prev;
local_reset_rise := resetBtn AND NOT reset_prev;

IF local_reset_rise THEN
    fillsToday := 0;
    local_accumVol := 0.0;
    valveOpen := FALSE;
    pendingConfirm := FALSE;
ELSE
    IF local_start_rise AND NOT valveOpen THEN
        local_accumVol := 0.0;
        valveOpen := TRUE;
        pendingConfirm := FALSE;
    END_IF;

    IF valveOpen THEN
        local_accumVol := local_accumVol + flowVol;
        IF local_accumVol >= targetVol THEN
            valveOpen := FALSE;
            pendingConfirm := TRUE;
        END_IF;
    END_IF;

    IF pendingConfirm AND doneSensor THEN
        IF fillsToday < INT#32767 THEN
            fillsToday := fillsToday + 1;
        END_IF;
        pendingConfirm := FALSE;
    END_IF;
END_IF;

start_prev := startBtn;
reset_prev := resetBtn;
END_FUNCTION_BLOCK

(* ---- self-medium-04.raw_candidate_01.st ---- *)
FUNCTION_BLOCK FB
VAR_INPUT
    startBtn : BOOL;
    resetBtn : BOOL;
    doneSensor : BOOL;
    targetVol : REAL;
    flowVol : REAL;
END_VAR
VAR_OUTPUT
    valveOpen : BOOL;
    fillsToday : INT;
END_VAR
VAR
    start_prev : BOOL := FALSE;
    reset_prev : BOOL := FALSE;
    pendingConfirm : BOOL := FALSE;
    local_accumVol : REAL := 0.0;
    local_start_rise : BOOL;
    local_reset_rise : BOOL;
END_VAR

(* ENGINEERING_CONTRACT
valveOpen: set on start_rise while previous output closed; hold while accumulated volume < targetVol;
            reset_rise priority closes immediately (S2,S5,S7,S8,S9).
pendingConfirm: set when accumulated volume reaches targetVol and valve closes; cleared by reset, new start,
            or confirmation after doneSensor = TRUE (Step4,S10,S13,S14).
fillsToday: +1 on pendingConfirm AND doneSensor, saturating at INT#32767; reset_rise sets 0;
            monotonic except reset (S1,S3,S4,S6,S14).
accumVol: REAL, mL; targetVol and flowVol REAL, mL; comparison uses >=.
*)
(* CONTRACT_RULES [] *)

local_start_rise := startBtn AND NOT start_prev;
local_reset_rise := resetBtn AND NOT reset_prev;

IF local_reset_rise THEN
    fillsToday := 0;
    local_accumVol := 0.0;
    valveOpen := FALSE;
    pendingConfirm := FALSE;
ELSE
    IF local_start_rise AND NOT valveOpen THEN
        local_accumVol := 0.0;
        valveOpen := TRUE;
        pendingConfirm := FALSE;
    END_IF;

    IF valveOpen THEN
        local_accumVol := local_accumVol + flowVol;
        IF local_accumVol >= targetVol THEN
            valveOpen := FALSE;
            pendingConfirm := TRUE;
        END_IF;
    END_IF;

    IF pendingConfirm AND doneSensor THEN
        IF fillsToday < INT#32767 THEN
            fillsToday := fillsToday + 1;
        END_IF;
        pendingConfirm := FALSE;
    END_IF;
END_IF;

start_prev := startBtn;
reset_prev := resetBtn;
END_FUNCTION_BLOCK

(* ---- self-medium-05.candidate_01.st ---- *)
(* ENGINEERING_CONTRACT
  qualified: combinational; TRUE when steamTemp in [447.0,453.0] and steamPressure in [3750.0,3850.0] (closed intervals) (PUB001,PUB004,S1).
  dataFault: combinational; TRUE when scanSeconds<=0 or >10, steamFlow<0 or >90, fuelFlow<0 or >6 (PUB003,PUB004,S4).
  qualifiedTon/fuelTon: retained accumulators; reset to 0 only on rising resetBtn; no accumulation on the reset scan (PUB004,PUB006,PUB007,S3,S9).
  With no reset edge and enable=TRUE and no dataFault: fuelTon increases; qualifiedTon increases only when qualified (PUB001,PUB002,PUB005,N10-S11,N10-S12).
  With no reset edge and enable=FALSE or dataFault=TRUE: accumulators hold their previous values (PUB006,S5,S6).
  revenue/cost/netProfit: recomputed every scan from current accumulators (PUB005,PUB008,S7).
  Units: flows kg/s, scanSeconds s, ton = kg/1000, revenue 280 CNY/t, cost 1500 CNY/t (PUB001,PUB008).
  resetBtn held TRUE after its edge does not repeatedly reset; only a new rising edge resets (PUB006,PUB007).
*)
(* CONTRACT_RULES [] *)
FUNCTION_BLOCK FB
VAR_INPUT
    enable : BOOL;
    resetBtn : BOOL;
    scanSeconds : LREAL;
    steamFlow : LREAL;
    fuelFlow : LREAL;
    steamTemp : LREAL;
    steamPressure : LREAL;
END_VAR
VAR_OUTPUT
    qualified : BOOL;
    dataFault : BOOL;
    qualifiedTon : LREAL;
    fuelTon : LREAL;
    revenue : LREAL;
    cost : LREAL;
    netProfit : LREAL;
END_VAR
VAR
    tmp_prev_reset : BOOL;
    tmp_reset_rise : BOOL;
    tmp_qualified_ton : LREAL;
    tmp_fuel_ton : LREAL;
END_VAR

    tmp_reset_rise := resetBtn AND NOT tmp_prev_reset;

    dataFault := (scanSeconds <= 0.0) OR (scanSeconds > 10.0)
                 OR (steamFlow < 0.0) OR (steamFlow > 90.0)
                 OR (fuelFlow < 0.0) OR (fuelFlow > 6.0);

    qualified := (steamTemp >= 447.0) AND (steamTemp <= 453.0)
                 AND (steamPressure >= 3750.0) AND (steamPressure <= 3850.0);

    IF tmp_reset_rise THEN
        tmp_qualified_ton := 0.0;
        tmp_fuel_ton := 0.0;
    ELSIF enable AND NOT dataFault THEN
        tmp_fuel_ton := tmp_fuel_ton + ((fuelFlow * scanSeconds) / 1000.0);
        IF qualified THEN
            tmp_qualified_ton := tmp_qualified_ton + ((steamFlow * scanSeconds) / 1000.0);
        END_IF;
    END_IF;

    tmp_prev_reset := resetBtn;

    qualifiedTon := tmp_qualified_ton;
    fuelTon := tmp_fuel_ton;
    revenue := tmp_qualified_ton * 280.0;
    cost := tmp_fuel_ton * 1500.0;
    netProfit := revenue - cost;

END_FUNCTION_BLOCK

(* ---- self-medium-05.raw_candidate_01.st ---- *)
(* ENGINEERING_CONTRACT
  qualified: combinational; TRUE when steamTemp in [447.0,453.0] and steamPressure in [3750.0,3850.0] (closed intervals) (PUB001,PUB004,S1).
  dataFault: combinational; TRUE when scanSeconds<=0 or >10, steamFlow<0 or >90, fuelFlow<0 or >6 (PUB003,PUB004,S4).
  qualifiedTon/fuelTon: retained accumulators; reset to 0 only on rising resetBtn; no accumulation on the reset scan (PUB004,PUB006,PUB007,S3,S9).
  With no reset edge and enable=TRUE and no dataFault: fuelTon increases; qualifiedTon increases only when qualified (PUB001,PUB002,PUB005,N10-S11,N10-S12).
  With no reset edge and enable=FALSE or dataFault=TRUE: accumulators hold their previous values (PUB006,S5,S6).
  revenue/cost/netProfit: recomputed every scan from current accumulators (PUB005,PUB008,S7).
  Units: flows kg/s, scanSeconds s, ton = kg/1000, revenue 280 CNY/t, cost 1500 CNY/t (PUB001,PUB008).
  resetBtn held TRUE after its edge does not repeatedly reset; only a new rising edge resets (PUB006,PUB007).
*)
(* CONTRACT_RULES [] *)
FUNCTION_BLOCK FB
VAR_INPUT
    enable : BOOL;
    resetBtn : BOOL;
    scanSeconds : LREAL;
    steamFlow : LREAL;
    fuelFlow : LREAL;
    steamTemp : LREAL;
    steamPressure : LREAL;
END_VAR
VAR_OUTPUT
    qualified : BOOL;
    dataFault : BOOL;
    qualifiedTon : LREAL;
    fuelTon : LREAL;
    revenue : LREAL;
    cost : LREAL;
    netProfit : LREAL;
END_VAR
VAR
    tmp_prev_reset : BOOL;
    tmp_reset_rise : BOOL;
    tmp_qualified_ton : LREAL;
    tmp_fuel_ton : LREAL;
END_VAR

    tmp_reset_rise := resetBtn AND NOT tmp_prev_reset;

    dataFault := (scanSeconds <= 0.0) OR (scanSeconds > 10.0)
                 OR (steamFlow < 0.0) OR (steamFlow > 90.0)
                 OR (fuelFlow < 0.0) OR (fuelFlow > 6.0);

    qualified := (steamTemp >= 447.0) AND (steamTemp <= 453.0)
                 AND (steamPressure >= 3750.0) AND (steamPressure <= 3850.0);

    IF tmp_reset_rise THEN
        tmp_qualified_ton := 0.0;
        tmp_fuel_ton := 0.0;
    ELSIF enable AND NOT dataFault THEN
        tmp_fuel_ton := tmp_fuel_ton + ((fuelFlow * scanSeconds) / 1000.0);
        IF qualified THEN
            tmp_qualified_ton := tmp_qualified_ton + ((steamFlow * scanSeconds) / 1000.0);
        END_IF;
    END_IF;

    tmp_prev_reset := resetBtn;

    qualifiedTon := tmp_qualified_ton;
    fuelTon := tmp_fuel_ton;
    revenue := tmp_qualified_ton * 280.0;
    cost := tmp_fuel_ton * 1500.0;
    netProfit := revenue - cost;

END_FUNCTION_BLOCK

(* ---- self-medium-06.candidate_01.st ---- *)
FUNCTION_BLOCK FB
VAR_INPUT
    enable : BOOL;
    resetBtn : BOOL;
    sensorValid : BOOL;
    setpoint : REAL;
    temperature : REAL;
    scanSeconds : REAL;
    bias : REAL;
END_VAR
VAR_OUTPUT
    power : REAL;
    correction : REAL;
    fault : BOOL;
END_VAR
VAR
    ePrev : REAL := 0.0;
    historyValid : BOOL := FALSE;
    local_prevReset : BOOL := FALSE;
    local_risingReset : BOOL;
    local_e : REAL;
    local_de : REAL;
    local_x : REAL;
    local_y : REAL;
END_VAR

(* ENGINEERING_CONTRACT
- power : computed via 20x+10y then clamped to [0,100]; zero when disabled/fault/reset rising. PUB001/PUB005/S1/S10/S11.
- correction : computed via 20x+10y, range [-30,30]; zero when disabled/fault/reset rising. PUB002/PUB004/S2.
- fault : combinational = NOT sensorValid OR scanSeconds<=0 OR scanSeconds>10; no retention. PUB003/S4/S5.
- historyValid/ePrev : cleared on disable/fault/reset rising; set after normal calculation; first/recovery scan uses de=0. PUB006/S7/S8/S12/S13.
- resetBtn edge : only rising edge triggers zero/clear; level hold does not keep zero. PUB009/S9.
- priority : fault/!enable/reset rising override normal calculation on same scan. PUB010/S3/S10.
- unspecified : NaN input behavior not specified; standard REAL LIMIT semantics used for clamps.
*)

(* CONTRACT_RULES [] *)

fault := (NOT sensorValid) OR (scanSeconds <= 0.0) OR (scanSeconds > 10.0);
local_risingReset := resetBtn AND NOT local_prevReset;

IF (NOT enable) OR fault OR local_risingReset THEN
    power := 0.0;
    correction := 0.0;
    ePrev := 0.0;
    historyValid := FALSE;
ELSE
    local_e := setpoint - temperature;

    IF NOT historyValid THEN
        local_de := 0.0;
    ELSE
        local_de := (local_e - ePrev) / scanSeconds;
    END_IF;

    local_x := LIMIT(-1.0, local_e / 10.0, 1.0);
    local_y := LIMIT(-1.0, local_de / 2.0, 1.0);

    correction := 20.0 * local_x + 10.0 * local_y;
    power := LIMIT(0.0, bias + correction, 100.0);

    ePrev := local_e;
    historyValid := TRUE;
END_IF;

local_prevReset := resetBtn;
END_FUNCTION_BLOCK

(* ---- self-medium-06.raw_candidate_01.st ---- *)
FUNCTION_BLOCK FB
VAR_INPUT
    enable : BOOL;
    resetBtn : BOOL;
    sensorValid : BOOL;
    setpoint : REAL;
    temperature : REAL;
    scanSeconds : REAL;
    bias : REAL;
END_VAR
VAR_OUTPUT
    power : REAL;
    correction : REAL;
    fault : BOOL;
END_VAR
VAR
    ePrev : REAL := 0.0;
    historyValid : BOOL := FALSE;
    local_prevReset : BOOL := FALSE;
    local_risingReset : BOOL;
    local_e : REAL;
    local_de : REAL;
    local_x : REAL;
    local_y : REAL;
END_VAR

(* ENGINEERING_CONTRACT
- power : computed via 20x+10y then clamped to [0,100]; zero when disabled/fault/reset rising. PUB001/PUB005/S1/S10/S11.
- correction : computed via 20x+10y, range [-30,30]; zero when disabled/fault/reset rising. PUB002/PUB004/S2.
- fault : combinational = NOT sensorValid OR scanSeconds<=0 OR scanSeconds>10; no retention. PUB003/S4/S5.
- historyValid/ePrev : cleared on disable/fault/reset rising; set after normal calculation; first/recovery scan uses de=0. PUB006/S7/S8/S12/S13.
- resetBtn edge : only rising edge triggers zero/clear; level hold does not keep zero. PUB009/S9.
- priority : fault/!enable/reset rising override normal calculation on same scan. PUB010/S3/S10.
- unspecified : NaN input behavior not specified; standard REAL LIMIT semantics used for clamps.
*)

(* CONTRACT_RULES [] *)

fault := (NOT sensorValid) OR (scanSeconds <= 0.0) OR (scanSeconds > 10.0);
local_risingReset := resetBtn AND NOT local_prevReset;

IF (NOT enable) OR fault OR local_risingReset THEN
    power := 0.0;
    correction := 0.0;
    ePrev := 0.0;
    historyValid := FALSE;
ELSE
    local_e := setpoint - temperature;

    IF NOT historyValid THEN
        local_de := 0.0;
    ELSE
        local_de := (local_e - ePrev) / scanSeconds;
    END_IF;

    local_x := LIMIT(-1.0, local_e / 10.0, 1.0);
    local_y := LIMIT(-1.0, local_de / 2.0, 1.0);

    correction := 20.0 * local_x + 10.0 * local_y;
    power := LIMIT(0.0, bias + correction, 100.0);

    ePrev := local_e;
    historyValid := TRUE;
END_IF;

local_prevReset := resetBtn;
END_FUNCTION_BLOCK
